            num nMoveType = 7
            num nPercentage
            num nSigValue
        pointRx pPointRx[2] = {x=278.890712, y=136.745171, z=230.948915, rx=84.337923, ry=-1.664851, rz=172.690172, shoulder=lefty, elbow=enegative, wrist=wnegative}
        string sID
      [1]
        bool bMarked
        jointRx jJointRx = {j1=14.463054, j2=126.686617, j3=-94.408556, j4=-18.307578, j5=-113.737208, j6=85.971215}
        pointRx pInter
        paraItem pParaItem
          [0]
            bool bSafePoint
            ifItem iIfItem
              [0]
                bool bANDOR[2]
                num nSigIndex[3]
                num nSigType[3]
                num nValue[3]
            mdesc mMdesc
            num nActionIndex = 71
            num nDelay = 1
            num nMoveType = 4
            num nPercentage
            num nSigValue
        pointRx pPointRx[2] = {x=278.890712, y=136.745171, z=230.948915, rx=84.337923, ry=-1.664851, rz=172.690172, shoulder=lefty, elbow=enegative, wrist=wnegative}
        string sID
      [2]
        bool bMarked
        jointRx jJointRx = {j1=14.463054, j2=126.686617, j3=-94.408556, j4=-18.307578, j5=-113.737208, j6=85.971215}
        pointRx pInter
        paraItem pParaItem
          [0]
            bool bSafePoint
            ifItem iIfItem
              [0]
                bool bANDOR[2]
                num nSigIndex[3]
                num nSigType[3]
                num nValue[3]
            mdesc mMdesc
            num nActionIndex = 70
            num nDelay = 1
            num nMoveType = 4
            num nPercentage
            num nSigValue = 1
        pointRx pPointRx[2] = {x=278.890712, y=136.745171, z=230.948915, rx=84.337923, ry=-1.664851, rz=172.690172, shoulder=lefty, elbow=enegative, wrist=wnegative}
        string sID
      [3]
        bool bMarked
        jointRx jJointRx = {j1=14.463054, j2=126.686617, j3=-94.408556, j4=-18.307578, j5=-113.737208, j6=85.971215}
        pointRx pInter
        paraItem pParaItem
          [0]
            bool bSafePoint
            ifItem iIfItem
              [0]
                bool bANDOR[2]
                num nSigIndex[3]
                num nSigType[3]
                num nValue[3]
            mdesc mMdesc
            num nActionIndex = 70
            num nDelay = 1
            num nMoveType = 3
            num nPercentage
            num nSigValue = 1
        pointRx pPointRx[2] = {x=278.890712, y=136.745171, z=230.948915, rx=84.337923, ry=-1.664851, rz=172.690172, shoulder=lefty, elbow=enegative, wrist=wnegative}
        string sID
      [4]
        bool bMarked
        jointRx jJointRx = {j1=-0.746077, j2=38.654193, j3=103.0610419, j4=-179.633028, j5=123.454226, j6=8.386419}
        pointRx pInter
        paraItem pParaItem
          [0]
            bool bSafePoint
            ifItem iIfItem
              [0]
                bool bANDOR[2]
                num nSigIndex[3]
                num nSigType[3]
                num nValue[3]
            mdesc mMdesc = {leave=0}
            num nActionIndex = 41
            num nDelay = 1
            num nMoveType = 1
            num nPercentage
            num nSigValue
        pointRx pPointRx[2] = {x=872.305806, y=193.820048, z=536.464849, rx=0.56853, ry=18.254398, rz=-172.702509, shoulder=lefty, elbow=epositive, wrist=wpositive}
        string sID
      [5]
        bool bMarked
        jointRx jJointRx = {j1=50.992067, j2=4.166676, j3=69.41419, j4=-184.312405, j5=69.584552, j6=-50.407158}
        pointRx pInter
        paraItem pParaItem
          [0]
            bool bSafePoint
            ifItem iIfItem
              [0]
                bool bANDOR[2]
                num nSigIndex[3]
                num nSigType[3]
                num nValue[3]
            mdesc mMdesc = {leave=0}
            num nActionIndex = 41
            num nDelay = 1
            num nMoveType = 1
            num nPercentage
            num nSigValue
        pointRx pPointRx[2] = {x=343.557382, y=727.163295, z=1235.32552, rx=-5.687342, ry=-0.597155, rz=179.191396, shoulder=lefty, elbow=epositive, wrist=wpositive}
        string sID
      [6]
        bool bMarked
        jointRx jJointRx = {j1=48.664808, j2=0.891331, j3=74.703897, j4=-185.753759, j5=70.406466, j6=-47.749335}
        pointRx pInter
        paraItem pParaItem
          [0]
            bool bSafePoint
            ifItem iIfItem
              [0]
                bool bANDOR[2]
                num nSigIndex[3]
                num nSigType[3]
                num nValue[3]
            mdesc mMdesc = {leave=0}
            num nActionIndex = 41
            num nDelay = 1
            num nMoveType = 1
            num nPercentage
            num nSigValue
        pointRx pPointRx[2] = {x=348.466857, y=713.703352, z=1210.583118, rx=-7.537716, ry=-0.596285, rz=179.191017, shoulder=lefty, elbow=epositive, wrist=wpositive}
        string sID
      [7]
        bool bMarked
        jointRx jJointRx = {j1=50.159419, j2=2.345991, j3=76.498933, j4=-185.508737, j5=73.496795, j6=-49.60951}
        pointRx pInter
        paraItem pParaItem
          [0]
            bool bSafePoint
            ifItem iIfItem
              [0]
                bool bANDOR[2]
                num nSigIndex[3]
                num nSigType[3]
                num nValue[3]
            mdesc mMdesc = {leave=0}
            num nActionIndex = 41
            num nDelay = 1
            num nMoveType = 1
            num nPercentage
            num nSigValue
        pointRx pPointRx[2] = {x=348.466871, y=737.786918, z=1179.801578, rx=-7.538916, ry=-0.596517, rz=179.191475, shoulder=lefty, elbow=epositive, wrist=wpositive}
        string sID
      [8]
        bool bMarked
        jointRx jJointRx = {j1=48.294816, j2=-0.682794, j3=80.800955, j4=-185.648441, j5=74.943082, j6=-47.842447}
        pointRx pInter
        paraItem pParaItem
          [0]
            bool bSafePoint
            ifItem iIfItem
              [0]
                bool bANDOR[2]
                num nSigIndex[3]
                num nSigType[3]
                num nValue[3]
            mdesc mMdesc = {leave=0}
            num nActionIndex = 41
            num nDelay = 1
            num nMoveType = 1
            num nPercentage
            num nSigValue
        pointRx pPointRx[2] = {x=348.466869, y=707.980912, z=1168.172739, rx=-7.537909, ry=-0.59668, rz=179.191275, shoulder=lefty, elbow=epositive, wrist=wpositive}
        string sID
      [9]
        bool bMarked
        jointRx jJointRx = {j1=59.661385, j2=20.184318, j3=65.0373942, j4=-180.17837, j5=86.0982717, j6=-60.460334}
        pointRx pInter
        paraItem pParaItem
          [0]
            bool bSafePoint
            ifItem iIfItem
              [0]
                bool bANDOR[2]
                num nSigIndex[3]
                num nSigType[3]
                num nValue[3]
            mdesc mMdesc = {leave=0}
            num nActionIndex = 41
            num nDelay = 1
            num nMoveType = 1
            num nPercentage
            num nSigValue
        pointRx pPointRx[2] = {x=342.103434, y=843.326292, z=1116.920644, rx=0.666634, ry=-0.596327, rz=179.191022, shoulder=lefty, elbow=epositive, wrist=wpositive}
        string sID
      [10]
        bool bMarked
        jointRx jJointRx = {j1=56.900837, j2=12.778869, j3=75.982676, j4=-180.135563, j5=89.64603, j6=-57.711316}
        pointRx pInter
        paraItem pParaItem
          [0]
            bool bSafePoint
            ifItem iIfItem
              [0]
                bool bANDOR[2]
                num nSigIndex[3]
                num nSigType[3]
                num nValue[3]
            mdesc mMdesc = {leave=0}
            num nActionIndex = 41
            num nDelay = 1
            num nMoveType = 1
            num nPercentage
            num nSigValue
        pointRx pPointRx[2] = {x=342.103419, y=775.469992, z=1101.315472, rx=0.666948, ry=-0.59656, rz=179.191109, shoulder=lefty, elbow=epositive, wrist=wpositive}
        string sID
      [11]
        bool bMarked
        jointRx jJointRx = {j1=56.518584, j2=13.362266, j3=64.344107, j4=-180.131909, j5=78.591486, j6=-57.304192}
        pointRx pInter
        paraItem pParaItem
          [0]
            bool bSafePoint
            ifItem iIfItem
              [0]
                bool bANDOR[2]
                num nSigIndex[3]
                num nSigType[3]
                num nValue[3]
            mdesc mMdesc = {leave=0}
            num nActionIndex = 41
            num nDelay = 1
            num nMoveType = 1
            num nPercentage
            num nSigValue
        pointRx pPointRx[2] = {x=342.103413, y=766.871901, z=1205.383601, rx=0.666905, ry=-0.596108, rz=179.190771, shoulder=lefty, elbow=epositive, wrist=wpositive}
        string sID
      [12]
        bool bMarked
        jointRx jJointRx = {j1=57.109214, j2=15.41659, j3=59.489821, j4=-180.142956, j5=75.789646, j6=-57.885688}
        pointRx pInter
        paraItem pParaItem
          [0]
            bool bSafePoint
            ifItem iIfItem
              [0]
                bool bANDOR[2]
                num nSigIndex[3]
                num nSigType[3]
                num nValue[3]
            mdesc mMdesc = {leave=0}
            num nActionIndex = 41
            num nDelay = 1
            num nMoveType = 1
            num nPercentage
            num nSigValue
        pointRx pPointRx[2] = {x=341.732761, y=779.650641, z=1227.038444, rx=0.666388, ry=-0.595966, rz=179.19083, shoulder=lefty, elbow=epositive, wrist=wpositive}
        string sID
      [13]
        bool bMarked
        jointRx jJointRx = {j1=39.164225, j2=-13.645288, j3=89.368263, j4=-186.463269, j5=70.113322, j6=-37.940152}
        pointRx pInter
        paraItem pParaItem
          [0]
            bool bSafePoint
            ifItem iIfItem
              [0]
                bool bANDOR[2]
                num nSigIndex[3]
                num nSigType[3]
                num nValue[3]
            mdesc mMdesc = {leave=0}
            num nActionIndex = 41
            num nDelay = 1
            num nMoveType = 1
            num nPercentage
            num nSigValue
        pointRx pPointRx[2] = {x=336.826434, y=577.61711, z=1191.998985, rx=-8.322487, ry=0.577625, rz=179.363473, shoulder=lefty, elbow=epositive, wrist=wpositive}
        string sID
      [14]
        bool bMarked
        jointRx jJointRx = {j1=32.650658, j2=-18.348971, j3=92.921174, j4=-187.128582, j5=69.716888, j6=-31.139541}
        pointRx pInter
        paraItem pParaItem
          [0]
            bool bSafePoint
            ifItem iIfItem
              [0]
                bool bANDOR[2]
                num nSigIndex[3]
                num nSigType[3]
                num nValue[3]
            mdesc mMdesc = {leave=0}
            num nActionIndex = 41
            num nDelay = 1
            num nMoveType = 1
            num nPercentage
            num nSigValue
        pointRx pPointRx[2] = {x=336.826433, y=515.325546, z=1191.37341, rx=-8.321046, ry=0.57803, rz=179.362899, shoulder=lefty, elbow=epositive, wrist=wpositive}
        string sID
      [15]
        bool bMarked
        jointRx jJointRx = {j1=36.0807313, j2=-9.953527, j3=74.825297, j4=-187.389169, j5=59.689212, j6=-33.315147}
        pointRx pInter
        paraItem pParaItem
          [0]
            bool bSafePoint
            ifItem iIfItem
              [0]
                bool bANDOR[2]
                num nSigIndex[3]
                num nSigType[3]
                num nValue[3]
            mdesc mMdesc = {leave=0}
            num nActionIndex = 41
            num nDelay = 1
            num nMoveType = 1
            num nPercentage
            num nSigValue
        pointRx pPointRx[2] = {x=351.37517, y=557.347514, z=1296.509025, rx=-8.32156, ry=0.577367, rz=179.363305, shoulder=lefty, elbow=epositive, wrist=wpositive}
        string sID
      [16]
        bool bMarked
        jointRx jJointRx = {j1=10.255909, j2=-18.0600505, j3=72.672032, j4=-190.141464, j5=52.980602, j6=-4.934383}
        pointRx pInter
        paraItem pParaItem
          [0]
            bool bSafePoint
            ifItem iIfItem
              [0]
                bool bANDOR[2]
                num nSigIndex[3]
                num nSigType[3]
                num nValue[3]
            mdesc mMdesc = {leave=0}
            num nActionIndex = 41
            num nDelay = 1
            num nMoveType = 1
            num nPercentage
            num nSigValue
        pointRx pPointRx[2] = {x=336.826448, y=355.459415, z=1364.362899, rx=-8.320098, ry=0.578249, rz=179.362643, shoulder=lefty, elbow=epositive, wrist=wpositive}
        string sID
      [17]
        bool bMarked
        jointRx jJointRx = {j1=90.161251, j2=-18.0722636, j3=77.256744, j4=-170.510373, j5=61.0400468, j6=-185.0917365}
        pointRx pInter
        paraItem pParaItem
          [0]
            bool bSafePoint
            ifItem iIfItem
              [0]
                bool bANDOR[2]
                num nSigIndex[3]
                num nSigType[3]
                num nValue[3]
            mdesc mMdesc = {leave=0}
            num nActionIndex = 41
            num nDelay = 1
            num nMoveType = 1
            num nPercentage
            num nSigValue
        pointRx pPointRx[2] = {x=193.885364, y=351.358286, z=1327.494019, rx=1.496376, ry=8.2983, rz=89.698418, shoulder=lefty, elbow=epositive, wrist=wpositive}
        string sID
      [18]
        bool bMarked
        jointRx jJointRx = {j1=76.262282, j2=-18.404812, j3=94.146484, j4=-169.188599, j5=85.00435766, j6=-167.549825}
        pointRx pInter
        paraItem pParaItem
          [0]
            bool bSafePoint
            ifItem iIfItem
              [0]
                bool bANDOR[2]
                num nSigIndex[3]
                num nSigType[3]
                num nValue[3]
            mdesc mMdesc = {leave=0}
            num nActionIndex = 41
            num nDelay = 1
            num nMoveType = 1
            num nPercentage
            num nSigValue
        pointRx pPointRx[2] = {x=297.323672, y=310.761188, z=1168.980461, rx=11.454003, ry=8.298378, rz=89.697972, shoulder=lefty, elbow=epositive, wrist=wpositive}
        string sID
      [19]
        bool bMarked
        jointRx jJointRx = {j1=126.372801, j2=0.947016, j3=58.247522, j4=-173.633502, j5=65.467797, j6=-219.528921}
        pointRx pInter
        paraItem pParaItem
          [0]
            bool bSafePoint
            ifItem iIfItem
              [0]
                bool bANDOR[2]
                num nSigIndex[3]
                num nSigType[3]
                num nValue[3]
            mdesc mMdesc = {leave=0}
            num nActionIndex = 41
            num nDelay = 1
            num nMoveType = 1
            num nPercentage
            num nSigValue
        pointRx pPointRx[2] = {x=-110.0468221, y=381.881454, z=1352.0109929, rx=1.496598, ry=8.298005, rz=89.698483, shoulder=lefty, elbow=epositive, wrist=wpositive}
        string sID
      [20]
        bool bMarked
        jointRx jJointRx = {j1=138.772753, j2=12.465275, j3=53.540842, j4=-175.467559, j5=73.29136, j6=-230.546088}
        pointRx pInter
        paraItem pParaItem
          [0]
            bool bSafePoint
            ifItem iIfItem
              [0]
                bool bANDOR[2]
                num nSigIndex[3]
                num nSigType[3]
                num nValue[3]
            mdesc mMdesc = {leave=0}
            num nActionIndex = 41
            num nDelay = 1
            num nMoveType = 1
            num nPercentage
            num nSigValue
        pointRx pPointRx[2] = {x=-284.713057, y=381.881445, z=1282.27146, rx=1.496715, ry=8.298986, rz=89.698256, shoulder=lefty, elbow=epositive, wrist=wpositive}
        string sID
      [21]
        bool bMarked
        jointRx jJointRx = {j1=129.569522, j2=-2.763661, j3=86.443161, j4=-174.560173, j5=90.131021, j6=-220.057051}
        pointRx pInter
        paraItem pParaItem
          [0]
            bool bSafePoint
            ifItem iIfItem
              [0]
                bool bANDOR[2]
                num nSigIndex[3]
                num nSigType[3]
                num nValue[3]
            mdesc mMdesc = {leave=0}
            num nActionIndex = 41
            num nDelay = 1
            num nMoveType = 1
            num nPercentage
            num nSigValue
        pointRx pPointRx[2] = {x=-158.339339, y=393.754355, z=1130.374707, rx=1.496575, ry=8.298917, rz=89.698258, shoulder=lefty, elbow=epositive, wrist=wpositive}
        string sID
      [22]
        bool bMarked
        jointRx jJointRx = {j1=141.483674, j2=14.580293, j3=86.0660414, j4=-182.560432, j5=99.634816, j6=-231.106968}
        pointRx pInter
        paraItem pParaItem
          [0]
            bool bSafePoint
            ifItem iIfItem
              [0]
                bool bANDOR[2]
                num nSigIndex[3]
                num nSigType[3]
                num nValue[3]
            mdesc mMdesc = {leave=0}
            num nActionIndex = 41
            num nDelay = 1
            num nMoveType = 1
            num nPercentage
            num nSigValue
        pointRx pPointRx[2] = {x=-456.482312, y=395.0927041, z=988.243024, rx=1.352323, ry=-2.355377, rz=90.855398, shoulder=lefty, elbow=epositive, wrist=wpositive}
        string sID
      [23]
        bool bMarked
        jointRx jJointRx = {j1=46.220955, j2=-26.278248, j3=73.480924, j4=-176.710401, j5=48.400229, j6=-56.2638}
        pointRx pInter
        paraItem pParaItem
          [0]
            bool bSafePoint
            ifItem iIfItem
              [0]
                bool bANDOR[2]
                num nSigIndex[3]
                num nSigType[3]
                num nValue[3]
            mdesc mMdesc = {leave=0}
            num nActionIndex = 41
            num nDelay = 1
            num nMoveType = 1
            num nPercentage
            num nSigValue
        pointRx pPointRx[2] = {x=156.67875, y=334.103919, z=1427.956714, rx=2.532212, ry=0.979884, rz=172.14558, shoulder=lefty, elbow=epositive, wrist=wpositive}
        string sID
      [24]
        bool bMarked
        jointRx jJointRx = {j1=-0.746077, j2=38.654193, j3=103.0610419, j4=-179.633028, j5=123.454226, j6=8.386419}
        pointRx pInter
        paraItem pParaItem
          [0]
            bool bSafePoint
            ifItem iIfItem
              [0]
                bool bANDOR[2]
                num nSigIndex[3]
                num nSigType[3]
                num nValue[3]
            mdesc mMdesc = {leave=10}
            num nActionIndex = 41
            num nDelay = 1
            num nMoveType = 1
            num nPercentage
            num nSigValue
        pointRx pPointRx[2] = {x=872.305806, y=193.820048, z=536.464849, rx=0.56853, ry=18.254398, rz=-172.702509, shoulder=lefty, elbow=epositive, wrist=wpositive}
        string sID
      [25]
        bool bMarked
        jointRx jJointRx = {j1=-0.746077, j2=38.654193, j3=103.0610419, j4=-179.633028, j5=123.454226, j6=8.386419}
        pointRx pInter
        paraItem pParaItem
          [0]
            bool bSafePoint
            ifItem iIfItem
              [0]
                bool bANDOR[2]
                num nSigIndex[3]
                num nSigType[3]
                num nValue[3]
            mdesc mMdesc = {leave=10}
            num nActionIndex = 70
            num nDelay = 1
            num nMoveType = 4
            num nPercentage
            num nSigValue
        pointRx pPointRx[2] = {x=872.305806, y=193.820048, z=536.464849, rx=0.56853, ry=18.254398, rz=-172.702509, shoulder=lefty, elbow=epositive, wrist=wpositive}
        string sID
      [26]
        bool bMarked
        jointRx jJointRx = {j1=-0.746077, j2=38.654193, j3=103.0610419, j4=-179.633028, j5=123.454226, j6=8.386419}
        pointRx pInter
        paraItem pParaItem
          [0]
            bool bSafePoint
            ifItem iIfItem
              [0]
                bool bANDOR[2]
                num nSigIndex[3]
                num nSigType[3]
                num nValue[3]
            mdesc mMdesc = {leave=10}
            num nActionIndex = 71
            num nDelay = 1
            num nMoveType = 4
            num nPercentage
            num nSigValue = 1
        pointRx pPointRx[2] = {x=872.305806, y=193.820048, z=536.464849, rx=0.56853, ry=18.254398, rz=-172.702509, shoulder=lefty, elbow=epositive, wrist=wpositive}
        string sID
      [27]
        bool bMarked
        jointRx jJointRx = {j1=-0.746077, j2=38.654193, j3=103.0610419, j4=-179.633028, j5=123.454226, j6=8.386419}
        pointRx pInter
        paraItem pParaItem
          [0]
            bool bSafePoint
            ifItem iIfItem
              [0]
                bool bANDOR[2]
                num nSigIndex[3]
                num nSigType[3]
                num nValue[3]
            mdesc mMdesc = {leave=10}
            num nActionIndex = 71
            num nDelay = 1
            num nMoveType = 3
            num nPercentage
            num nSigValue = 1
        pointRx pPointRx[2] = {x=872.305806, y=193.820048, z=536.464849, rx=0.56853, ry=18.254398, rz=-172.702509, shoulder=lefty, elbow=epositive, wrist=wpositive}
        string sID
      [28]
        bool bMarked
        jointRx jJointRx = {j1=94.696904, j2=-17.194257, j3=77.457422, j4=-178.674473, j5=60.986606, j6=84.00973218}
        pointRx pInter
        paraItem pParaItem
          [0]
            bool bSafePoint
            ifItem iIfItem
              [0]
                bool bANDOR[2]
                num nSigIndex[3]
                num nSigType[3]
                num nValue[3]
            mdesc mMdesc = {leave=0}
            num nActionIndex = 41
            num nDelay = 1
            num nMoveType = 1
            num nPercentage
            num nSigValue
        pointRx pPointRx[2] = {x=-70.0312062, y=207.928659, z=1348.60192, rx=0.619605, ry=1.21397, rz=-0.649688, shoulder=lefty, elbow=epositive, wrist=wpositive}
        string sID
      [29]
        bool bMarked
        jointRx jJointRx = {j1=92.713698, j2=17.804684, j3=59.507036, j4=-178.795122, j5=71.278521, j6=86.0690239}
        pointRx pInter
        paraItem pParaItem
          [0]
            bool bSafePoint
            ifItem iIfItem
              [0]
                bool bANDOR[2]
                num nSigIndex[3]
                num nSigType[3]
                num nValue[3]
            mdesc mMdesc = {leave=0}
            num nActionIndex = 41
            num nDelay = 1
            num nMoveType = 1
            num nPercentage
            num nSigValue
        pointRx pPointRx[2] = {x=-78.365141, y=640.766438, z=1210.403131, rx=-6.0840607, ry=0.854555, rz=-0.845261, shoulder=lefty, elbow=epositive, wrist=wpositive}
        string sID
      [30]
        bool bMarked
        jointRx jJointRx = {j1=92.713698, j2=17.804684, j3=59.507036, j4=-178.795122, j5=71.278521, j6=86.0690239}
        pointRx pInter
        paraItem pParaItem
          [0]
            bool bSafePoint
            ifItem iIfItem
              [0]
                bool bANDOR[2]
                num nSigIndex[3]
                num nSigType[3]
                num nValue[3]
            mdesc mMdesc = {leave=0}
            num nActionIndex = 41
            num nDelay = 1
            num nMoveType = 7
            num nPercentage
            num nSigValue
        pointRx pPointRx[2] = {x=-78.365141, y=640.766438, z=1210.403131, rx=-6.0840607, ry=0.854555, rz=-0.845261, shoulder=lefty, elbow=epositive, wrist=wpositive}
        string sID
      [31]
        bool bMarked
        jointRx jJointRx = {j1=93.634054, j2=-0.200585, j3=81.614575, j4=-178.59677, j5=73.693191, j6=85.159231}
        pointRx pInter
        paraItem pParaItem
          [0]
            bool bSafePoint
            ifItem iIfItem
              [0]
                bool bANDOR[2]
                num nSigIndex[3]
                num nSigType[3]
                num nValue[3]
            mdesc mMdesc = {leave=0}
            num nActionIndex = 41
            num nDelay = 1
            num nMoveType = 1
            num nPercentage
            num nSigValue
        pointRx pPointRx[2] = {x=-80.825264, y=510.591299, z=1198.230863, rx=-7.794676, ry=0.855921, rz=-0.845268, shoulder=lefty, elbow=epositive, wrist=wpositive}
        string sID
      [32]
        bool bMarked
        jointRx jJointRx = {j1=93.634054, j2=-0.200585, j3=81.614575, j4=-178.59677, j5=73.693191, j6=85.159231}
        pointRx pInter
        paraItem pParaItem
          [0]
            bool bSafePoint
            ifItem iIfItem
              [0]
                bool bANDOR[2]
                num nSigIndex[3]
                num nSigType[3]
                num nValue[3]
            mdesc mMdesc = {leave=0}
            num nActionIndex = 41
            num nDelay = 1
            num nMoveType = 7
            num nPercentage
            num nSigValue
        pointRx pPointRx[2] = {x=-80.825264, y=510.591299, z=1198.230863, rx=-7.794676, ry=0.855921, rz=-0.845268, shoulder=lefty, elbow=epositive, wrist=wpositive}
        string sID
      [33]
        bool bMarked
        jointRx jJointRx = {j1=94.697022, j2=-26.101782, j3=117.801323, j4=-178.839759, j5=92.416802, j6=84.701619}
        pointRx pInter
        paraItem pParaItem
          [0]
            bool bSafePoint
            ifItem iIfItem
              [0]
                bool bANDOR[2]
                num nSigIndex[3]
                num nSigType[3]
                num nValue[3]
            mdesc mMdesc = {leave=0}
            num nActionIndex = 41
            num nDelay = 1
            num nMoveType = 1
            num nPercentage
            num nSigValue
        pointRx pPointRx[2] = {x=-70.0312042, y=207.928608, z=1030.831107, rx=0.620415, ry=1.214089, rz=-0.649604, shoulder=lefty, elbow=epositive, wrist=wpositive}
        string sID
      [34]
        bool bMarked
        jointRx jJointRx = {j1=-0.746077, j2=38.654194, j3=103.0610414, j4=-179.633029, j5=123.454226, j6=8.386419}
        pointRx pInter
        paraItem pParaItem
          [0]
            bool bSafePoint
            ifItem iIfItem
              [0]
                bool bANDOR[2]
                num nSigIndex[3]
                num nSigType[3]
                num nValue[3]
            mdesc mMdesc = {leave=0}
            num nActionIndex = 41
            num nDelay = 1
            num nMoveType = 1
            num nPercentage
            num nSigValue
        pointRx pPointRx[2] = {x=872.305806, y=193.820048, z=536.464849, rx=0.56853, ry=18.254398, rz=-172.702509, shoulder=lefty, elbow=epositive, wrist=wpositive}
        string sID
      [35]
        bool bMarked
        jointRx jJointRx = {j1=-0.746077, j2=38.654194, j3=103.0610414, j4=-179.633029, j5=123.454226, j6=8.386419}
        pointRx pInter
        paraItem pParaItem
          [0]
            bool bSafePoint
            ifItem iIfItem
              [0]
                bool bANDOR[2]
                num nSigIndex[3]
                num nSigType[3]
                num nValue[3]
            mdesc mMdesc = {leave=0}
            num nActionIndex = 71
            num nDelay = 1
            num nMoveType = 4
            num nPercentage
            num nSigValue
        pointRx pPointRx[2] = {x=872.305806, y=193.820048, z=536.464849, rx=0.56853, ry=18.254398, rz=-172.702509, shoulder=lefty, elbow=epositive, wrist=wpositive}
        string sID
      [36]
        bool bMarked
        jointRx jJointRx = {j1=-0.746077, j2=38.654194, j3=103.0610414, j4=-179.633029, j5=123.454226, j6=8.386419}
        pointRx pInter
        paraItem pParaItem
          [0]
            bool bSafePoint
            ifItem iIfItem
              [0]
                bool bANDOR[2]
                num nSigIndex[3]
                num nSigType[3]
                num nValue[3]
            mdesc mMdesc = {leave=0}
            num nActionIndex = 70
            num nDelay = 1
            num nMoveType = 4
            num nPercentage
            num nSigValue = 1
        pointRx pPointRx[2] = {x=872.305806, y=193.820048, z=536.464849, rx=0.56853, ry=18.254398, rz=-172.702509, shoulder=lefty, elbow=epositive, wrist=wpositive}
        string sID
      [37]
        bool bMarked
        jointRx jJointRx = {j1=-0.746077, j2=38.654194, j3=103.0610414, j4=-179.633029, j5=123.454226, j6=8.386419}
        pointRx pInter
        paraItem pParaItem
          [0]
            bool bSafePoint
            ifItem iIfItem
              [0]
                bool bANDOR[2]
                num nSigIndex[3]
                num nSigType[3]
                num nValue[3]
            mdesc mMdesc = {leave=0}
            num nActionIndex = 70
            num nDelay = 1
            num nMoveType = 3
            num nPercentage
            num nSigValue = 1
        pointRx pPointRx[2] = {x=872.305806, y=193.820048, z=536.464849, rx=0.56853, ry=18.254398, rz=-172.702509, shoulder=lefty, elbow=epositive, wrist=wpositive}
        string sID
    string sID
  [PR01_WashPath01]
    num nFrameIndex
    num nMoveID
    num nToolIndex
    pointItem pPointItem
      [0]
        bool bMarked
        jointRx jJointRx
        pointRx pInter
        paraItem pParaItem
          [0]
            bool bSafePoint
            ifItem iIfItem
              [0]
                bool bANDOR[2]
                num nSigIndex[3]
                num nSigType[3]
                num nValue[3]
            mdesc mMdesc
            num nActionIndex
            num nDelay
            num nMoveType
            num nPercentage
            num nSigValue
        pointRx pPointRx[2]
        string sID
    string sID
  [PR02-WashPATH1]
    num nFrameIndex
    num nMoveID
    num nToolIndex
    pointItem pPointItem[31]
      [0]
        bool bMarked
        jointRx jJointRx = {j1=14.463054, j2=126.686617, j3=-94.408556, j4=-18.307578, j5=-113.737208, j6=85.971215}
        pointRx pInter
        paraItem pParaItem
          [0]
            bool bSafePoint
            ifItem iIfItem
              [0]
                bool bANDOR[2]
                num nSigIndex[3]
                num nSigType[3]
                num nValue[3]
            mdesc mMdesc
            num nActionIndex = 41
            num nDelay = 1
            num nMoveType = 7
            num nPercentage
            num nSigValue
        pointRx pPointRx[2] = {x=278.890712, y=136.745171, z=230.948915, rx=84.337923, ry=-1.664851, rz=172.690172, shoulder=lefty, elbow=enegative, wrist=wnegative}
        string sID
      [1]
        bool bMarked
        jointRx jJointRx = {j1=14.463054, j2=126.686617, j3=-94.408556, j4=-18.307578, j5=-113.737208, j6=85.971215}
        pointRx pInter
        paraItem pParaItem
          [0]
            bool bSafePoint
            ifItem iIfItem
              [0]
                bool bANDOR[2]
                num nSigIndex[3]
                num nSigType[3]
                num nValue[3]
            mdesc mMdesc
            num nActionIndex = 71
            num nDelay = 1
            num nMoveType = 4
            num nPercentage
            num nSigValue
        pointRx pPointRx[2] = {x=278.890712, y=136.745171, z=230.948915, rx=84.337923, ry=-1.664851, rz=172.690172, shoulder=lefty, elbow=enegative, wrist=wnegative}
        string sID
      [2]
        bool bMarked
        jointRx jJointRx = {j1=14.463054, j2=126.686617, j3=-94.408556, j4=-18.307578, j5=-113.737208, j6=85.971215}
        pointRx pInter
        paraItem pParaItem
          [0]
            bool bSafePoint
            ifItem iIfItem
              [0]
                bool bANDOR[2]
                num nSigIndex[3]
                num nSigType[3]
                num nValue[3]
            mdesc mMdesc
            num nActionIndex = 70
            num nDelay = 1
            num nMoveType = 4
            num nPercentage
            num nSigValue = 1
        pointRx pPointRx[2] = {x=278.890712, y=136.745171, z=230.948915, rx=84.337923, ry=-1.664851, rz=172.690172, shoulder=lefty, elbow=enegative, wrist=wnegative}
        string sID
      [3]
        bool bMarked
        jointRx jJointRx = {j1=14.463054, j2=126.686617, j3=-94.408556, j4=-18.307578, j5=-113.737208, j6=85.971215}
        pointRx pInter
        paraItem pParaItem
          [0]
            bool bSafePoint
            ifItem iIfItem
              [0]
                bool bANDOR[2]
                num nSigIndex[3]
                num nSigType[3]
                num nValue[3]
            mdesc mMdesc
            num nActionIndex = 70
            num nDelay = 1
            num nMoveType = 3
            num nPercentage
            num nSigValue = 1
        pointRx pPointRx[2] = {x=278.890712, y=136.745171, z=230.948915, rx=84.337923, ry=-1.664851, rz=172.690172, shoulder=lefty, elbow=enegative, wrist=wnegative}
        string sID
      [4]
        bool bMarked
        jointRx jJointRx = {j1=-0.746077, j2=38.654193, j3=103.0610419, j4=-179.633028, j5=123.454226, j6=8.386419}
        pointRx pInter
        paraItem pParaItem
          [0]
            bool bSafePoint
            ifItem iIfItem
              [0]
                bool bANDOR[2]
                num nSigIndex[3]
                num nSigType[3]
                num nValue[3]
            mdesc mMdesc = {leave=0}
            num nActionIndex = 41
            num nDelay = 1
            num nMoveType = 1
            num nPercentage
            num nSigValue
        pointRx pPointRx[2] = {x=872.305806, y=193.820048, z=536.464849, rx=0.56853, ry=18.254398, rz=-172.702509, shoulder=lefty, elbow=epositive, wrist=wpositive}
        string sID
      [5]
        bool bMarked
        jointRx jJointRx = {j1=54.199422, j2=12.224855, j3=66.41542, j4=-178.0531166, j5=78.997815, j6=-52.670521}
        pointRx pInter
        paraItem pParaItem
          [0]
            bool bSafePoint
            ifItem iIfItem
              [0]
                bool bANDOR[2]
                num nSigIndex[3]
                num nSigType[3]
                num nValue[3]
            mdesc mMdesc = {leave=0}
            num nActionIndex = 41
            num nDelay = 1
            num nMoveType = 1
            num nPercentage
            num nSigValue
        pointRx pPointRx[2] = {x=374.858876, y=738.189444, z=1200.688847, rx=1.403036, ry=1.344431, rz=-178.110008, shoulder=lefty, elbow=epositive, wrist=wpositive}
        string sID
      [6]
        bool bMarked
        jointRx jJointRx = {j1=55.0834751, j2=13.697298, j3=67.00047558, j4=-178.0711603, j5=81.0838955, j6=-53.48245}
        pointRx pInter
        paraItem pParaItem
          [0]
            bool bSafePoint
            ifItem iIfItem
              [0]
                bool bANDOR[2]
                num nSigIndex[3]
                num nSigType[3]
                num nValue[3]
            mdesc mMdesc = {leave=0}
            num nActionIndex = 41
            num nDelay = 1
            num nMoveType = 1
            num nPercentage
            num nSigValue
        pointRx pPointRx[2] = {x=374.858872, y=756.93507, z=1178.378474, rx=1.403375, ry=1.344299, rz=-178.110043, shoulder=lefty, elbow=epositive, wrist=wpositive}
        string sID
      [7]
        bool bMarked
        jointRx jJointRx = {j1=50.804516, j2=5.425514, j3=70.291644, j4=-178.0123323, j5=75.962597, j6=-49.384227}
        pointRx pInter
        paraItem pParaItem
          [0]
            bool bSafePoint
            ifItem iIfItem
              [0]
                bool bANDOR[2]
                num nSigIndex[3]
                num nSigType[3]
                num nValue[3]
            mdesc mMdesc = {leave=0}
            num nActionIndex = 41
            num nDelay = 1
            num nMoveType = 1
            num nPercentage
            num nSigValue
        pointRx pPointRx[2] = {x=368.36511, y=665.236172, z=1237.143339, rx=1.402732, ry=1.344359, rz=-178.109873, shoulder=lefty, elbow=epositive, wrist=wpositive}
        string sID
      [8]
        bool bMarked
        jointRx jJointRx = {j1=45.633733, j2=4.768064, j3=58.245369, j4=-177.822903, j5=63.0908471, j6=-44.713841}
        pointRx pInter
        paraItem pParaItem
          [0]
            bool bSafePoint
            ifItem iIfItem
              [0]
                bool bANDOR[2]
                num nSigIndex[3]
                num nSigType[3]
